// TIA Portal V20 export
// export: Created 2026-10-19T18:06:28.1377235Z, ExportSetting WithDefaults, DisplayName Totally Integrated Automation Portal, DisplayVersion V20 Update 6, DisplayName TIA Portal Openness, DisplayVersion V20 Update 6, DisplayName TIA Portal Version Control Interface, DisplayVersion V20 Update 6, DisplayName SINAMICS Startdrive Advanced, DisplayVersion V20 SP1, DisplayName SINAMICS Startdrive G130, G150, S120, S150, SINAMICS MV, G220, S200, S210, DisplayVersion V20 SP1, DisplayName SINAMICS Startdrive G110M, G120, G120C, G120D, G120P, G115D, DisplayVersion V20 SP1, DisplayName STEP 7 Professional, DisplayVersion V20 Update 6, DisplayName STEP 7 Safety, DisplayVersion V20 Update 2, DisplayName WinCC Basic/Comfort/Advanced, DisplayVersion V20 Update 6, DisplayName WinCC Unified, DisplayVersion V20 Update 6
FUNCTION_BLOCK "SAI_IND_WriteAdjustSettings"   // FB51, LAD
{ S7_Optimized_Access := 'FALSE' }
VERSION : 0.1
// stored: AutoNumber true, IsIECCheckEnabled false, SetENOAutomatically false, UDAEnableTagReadback false
   VAR_INPUT
      ID : HW_IO;   // The Profinet Device Hardware Identifier under device properties
      ScaleCapacity : Real;   // Scale capacity to be written into the transmitter
      Increment : Real;   // Increment value to be written into the transmitter
   END_VAR
   VAR_OUTPUT
      Done : Bool;   // Write process done successfully
      Error : Bool;   // Error during writing process
   END_VAR
   VAR_IN_OUT
      Write : Bool;   // Switch this bit ON to start writing
   END_VAR
   VAR DB_SPECIFIC
      Static01 : Bool;
      "Step" : Int;
   END_VAR
   VAR
      WRREC_CAP { S7_SetPoint := 'True'} : WRREC;
   END_VAR
   VAR DB_SPECIFIC
      CAP_RECORD : Real;
      INC_RECORD : Real;
      Activate : Bool;
   END_VAR
   VAR_TEMP   // added for the SCL form of the ladder/FBD networks
      _w1 : Bool;
      _w2 : Bool;
      _w3 : Bool;
      _w4 : Bool;
      _w5 : Bool;
      _w6 : Bool;
      _w7 : Bool;
   END_VAR
BEGIN

REGION Network 1: Initialization and Checking
   // Initializes FB output bits:
   // Process;
   // Error;
   // Done;
   // Check validity of scale capacity and increment values before proceeding to next step
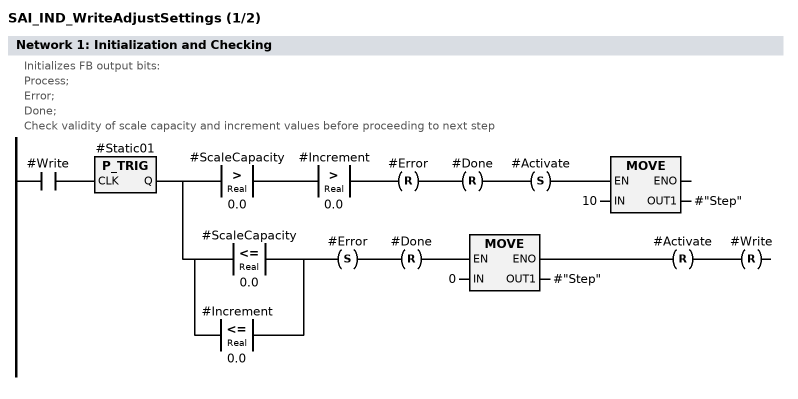
   RUNG wire#powerrail
      Contact( #Write )
      P_Trig( #Static01 )
      wire#w1
      { S7_Templates := "SrcType := Real" } GT_Contact(in1 := #ScaleCapacity, in2 := 0.0)
      { S7_Templates := "SrcType := Real" } GT_Contact(in1 := #Increment, in2 := 0.0)
      R_Coil( #Error )
      R_Coil( #Done )
      S_Coil( #Activate )
      { S7_GenerateENO := "TRUE" } Move(in := 10, out1 => #"Step")
   END_RUNG
   RUNG wire#w1
      { S7_Templates := "SrcType := Real" } LE_Contact(in1 := #ScaleCapacity, in2 := 0.0)
      wire#w2
      S_Coil( #Error )
      R_Coil( #Done )
      { S7_GenerateENO := "TRUE" } Move(in := 0, out1 => #"Step")
      R_Coil( #Activate )
      R_Coil( #Write )
   END_RUNG
   RUNG wire#w1
      { S7_Templates := "SrcType := Real" } LE_Contact(in1 := #Increment, in2 := 0.0)
   END_RUNG wire#w2
   // the same network as SCL:
   // ENO of a box is taken as its EN; it also drops when the box reports an error
   #_w1 := #Write AND NOT #Static01;   // rising edge
   #Static01 := #Write;
   IF #_w1 AND (#ScaleCapacity > 0.0) AND (#Increment > 0.0) THEN
       #Error := FALSE;
       #Done := FALSE;
       #Activate := TRUE;
       #"Step" := 10;
   END_IF;
   IF #_w1 AND ((#ScaleCapacity <= 0.0) OR (#Increment <= 0.0)) THEN
       #Error := TRUE;
       #Done := FALSE;
       #"Step" := 0;
       #Activate := FALSE;
       #Write := FALSE;
   END_IF;
END_REGION

REGION Network 2: Sequence
   // Sequence steps:
   // 10: Write in scale capacity (REAL; Index= 16#4367)
   // 20: Write in scale increment (REAL; Index= 16#4366)
   // 30: Completed the write process, DONE bit is set to TRUE
   // 99: ERROR bit is set to TRUE due to error
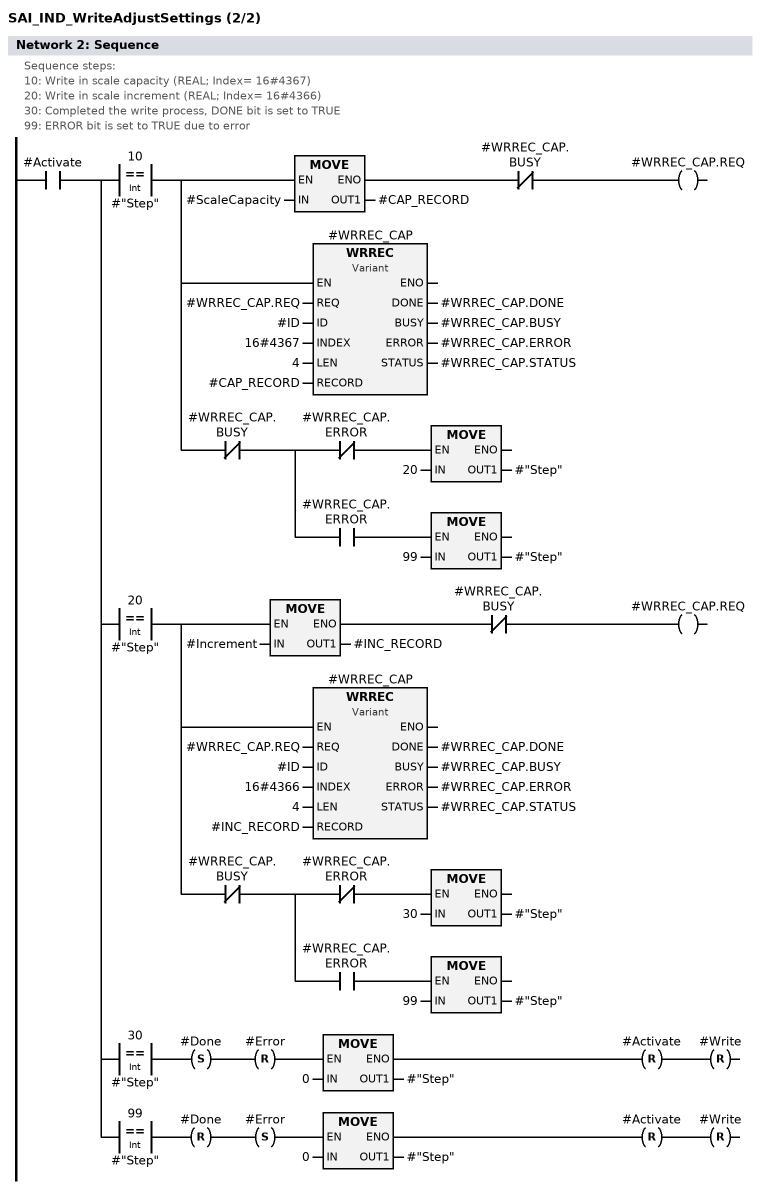
   RUNG wire#powerrail
      Contact( #Activate )
      wire#w1
      { S7_Templates := "SrcType := Int" } EQ_Contact(in1 := 10, in2 := #"Step")
      wire#w2
      { S7_GenerateENO := "TRUE" } Move(in := #ScaleCapacity, out1 => #CAP_RECORD)
      I_Contact( #WRREC_CAP.BUSY )
      Coil( #WRREC_CAP.REQ )
   END_RUNG
   RUNG wire#w2
      { S7_Templates := "[ptr_type := Variant, id_type := HW_IO, index_type := DInt, len_type := UInt]" } #WRREC_CAP.WRREC(REQ := #WRREC_CAP.REQ, ID := #ID, INDEX := 16#4367, LEN := 4, RECORD := #CAP_RECORD, DONE => #WRREC_CAP.DONE, BUSY => #WRREC_CAP.BUSY, ERROR => #WRREC_CAP.ERROR, STATUS => #WRREC_CAP.STATUS)
   END_RUNG
   RUNG wire#w2
      I_Contact( #WRREC_CAP.BUSY )
      wire#w3
      I_Contact( #WRREC_CAP.ERROR )
      { S7_GenerateENO := "TRUE" } Move(in := 20, out1 => #"Step")
   END_RUNG
   RUNG wire#w3
      Contact( #WRREC_CAP.ERROR )
      { S7_GenerateENO := "TRUE" } Move(in := 99, out1 => #"Step")
   END_RUNG
   RUNG wire#w1
      { S7_Templates := "SrcType := Int" } EQ_Contact(in1 := 20, in2 := #"Step")
      wire#w4
      { S7_GenerateENO := "TRUE" } Move(in := #Increment, out1 => #INC_RECORD)
      I_Contact( #WRREC_CAP.BUSY )
      Coil( #WRREC_CAP.REQ )
   END_RUNG
   RUNG wire#w4
      { S7_Templates := "[ptr_type := Variant, id_type := HW_IO, index_type := DInt, len_type := UInt]" } #WRREC_CAP.WRREC(REQ := #WRREC_CAP.REQ, ID := #ID, INDEX := 16#4366, LEN := 4, RECORD := #INC_RECORD, DONE => #WRREC_CAP.DONE, BUSY => #WRREC_CAP.BUSY, ERROR => #WRREC_CAP.ERROR, STATUS => #WRREC_CAP.STATUS)
   END_RUNG
   RUNG wire#w4
      I_Contact( #WRREC_CAP.BUSY )
      wire#w5
      I_Contact( #WRREC_CAP.ERROR )
      { S7_GenerateENO := "TRUE" } Move(in := 30, out1 => #"Step")
   END_RUNG
   RUNG wire#w5
      Contact( #WRREC_CAP.ERROR )
      { S7_GenerateENO := "TRUE" } Move(in := 99, out1 => #"Step")
   END_RUNG
   RUNG wire#w1
      { S7_Templates := "SrcType := Int" } EQ_Contact(in1 := 30, in2 := #"Step")
      S_Coil( #Done )
      R_Coil( #Error )
      { S7_GenerateENO := "TRUE" } Move(in := 0, out1 => #"Step")
      R_Coil( #Activate )
      R_Coil( #Write )
   END_RUNG
   RUNG wire#w1
      { S7_Templates := "SrcType := Int" } EQ_Contact(in1 := 99, in2 := #"Step")
      R_Coil( #Done )
      S_Coil( #Error )
      { S7_GenerateENO := "TRUE" } Move(in := 0, out1 => #"Step")
      R_Coil( #Activate )
      R_Coil( #Write )
   END_RUNG
   // the same network as SCL:
   // ENO of a box is taken as its EN; it also drops when the box reports an error
   #_w1 := #Activate AND (10 = #"Step");
   IF #_w1 THEN #CAP_RECORD := #ScaleCapacity; END_IF;
   #WRREC_CAP.REQ := #_w1 AND NOT #WRREC_CAP.BUSY;
   IF #_w1 THEN
       #WRREC_CAP(REQ := #WRREC_CAP.REQ,   // WRREC
                  ID := #ID,
                  INDEX := 16#4367,
                  LEN := 4,
                  RECORD := #CAP_RECORD,
                  DONE => #WRREC_CAP.DONE,
                  BUSY => #WRREC_CAP.BUSY,
                  ERROR => #WRREC_CAP.ERROR,
                  STATUS => #WRREC_CAP.STATUS);
   END_IF;
   #_w2 := #_w1 AND NOT #WRREC_CAP.BUSY;
   IF #_w2 AND NOT #WRREC_CAP.ERROR THEN #"Step" := 20; END_IF;
   IF #_w2 AND #WRREC_CAP.ERROR THEN #"Step" := 99; END_IF;
   #_w3 := #Activate AND (20 = #"Step");
   IF #_w3 THEN #INC_RECORD := #Increment; END_IF;
   #WRREC_CAP.REQ := #_w3 AND NOT #WRREC_CAP.BUSY;
   IF #_w3 THEN
       #WRREC_CAP(REQ := #WRREC_CAP.REQ,   // WRREC
                  ID := #ID,
                  INDEX := 16#4366,
                  LEN := 4,
                  RECORD := #INC_RECORD,
                  DONE => #WRREC_CAP.DONE,
                  BUSY => #WRREC_CAP.BUSY,
                  ERROR => #WRREC_CAP.ERROR,
                  STATUS => #WRREC_CAP.STATUS);
   END_IF;
   #_w4 := #_w3 AND NOT #WRREC_CAP.BUSY;
   IF #_w4 AND NOT #WRREC_CAP.ERROR THEN #"Step" := 30; END_IF;
   IF #_w4 AND #WRREC_CAP.ERROR THEN #"Step" := 99; END_IF;
   IF #Activate AND (30 = #"Step") THEN
       #Done := TRUE;
       #Error := FALSE;
   END_IF;
   #_w5 := #Activate AND (30 = #"Step");
   IF #_w5 THEN #"Step" := 0; END_IF;
   #_w6 := #Activate;
   IF #_w5 THEN
       #Activate := FALSE;
       #Write := FALSE;
   END_IF;
   IF #_w6 AND (99 = #"Step") THEN
       #Done := FALSE;
       #Error := TRUE;
   END_IF;
   #_w7 := #_w6 AND (99 = #"Step");
   IF #_w7 THEN
       #"Step" := 0;
       #Activate := FALSE;
       #Write := FALSE;
   END_IF;
END_REGION
END_FUNCTION_BLOCK
